(* EMS UPS 명령 1건 (MqttTask → PlcTask 칸, GVL_IF.g_astUpsCmd). 2026-11-05. 명세: WR-UPS-01 *)
TYPE ST_IfUpsCmd :
STRUCT
	nSeq	: UDINT;	// 새 명령마다 1씩 오름. 받는 쪽은 번호 변화로 새 명령을 안다
	nType	: UDINT;	// 명령 번호 1~26, 101 수동·102 자동 (EMS CommandType 그대로. 인터페이스 100.Command, 명세 WR-UPS-01)
END_STRUCT
END_TYPE

(* stored: Version 1.1.0.1, ProductVersion 3.1.4024.12
   DUT ST_IfUpsCmd: Id {cd5c9362-7f9b-4b8f-9584-eef02043a399} *)
